(* IEC 61131-3 sources: s7-to-codesys/s7conv/tests/snapshots/fixtures/src/POUs/FB_Legacy, 2 files *)

(* ---- FB_Legacy.decl.st ---- *)
// Назначение: Функциональный блок «FB_Legacy», сконвертирован из SCL
// Автор:      не указан (исходный блок S7); перевод в ST — s7conv 0.1.0
// Версия:     0.1 (исходный блок S7)
// Документ:   docs/CONVERSION_REPORT.md, docs/MAPPING.md
// Источник:   s7conv/tests/fixtures/unsupported.scl, строки 2–44, FUNCTION_BLOCK "FB_Legacy"
// Сгенерировано s7conv: пометки MIGRATION-CHECK и MIGRATION-TODO требуют ручного разбора.
// MIGRATION-CHECK: стандартный (неоптимизированный) доступ S7: абсолютная адресация и порядок байтов не переносятся
//                  (стр. 2)
// MIGRATION-CHECK: реманентность задаётся в экземпляре DB (DB_SPECIFIC) — объявлено VAR (стр. 19)
// ---- комментарий в начале исходного файла SCL ----
// Фикстура s7conv: конструкции, которые конвертер не переводит или переводит с пометкой.
FUNCTION_BLOCK FB_Legacy
VAR_INPUT
    // MIGRATION-TODO: Variant — нет аналога в CODESYS; переписать (ANY, POINTER или перегрузка) (стр. 6)
    // anyIn : Variant;
    // MIGRATION-TODO: DTL — структура S7 (YEAR, MONTH, ...), в CODESYS нет; заменить на DT или свою структуру (стр.
    //                 7)
    // stamp : DTL;
    // MIGRATION-CHECK: имя «time» переименовано в «time_» (ключевое слово CODESYS или повтор) (стр. 8)
    time_ : TIME;
END_VAR
VAR
    raw : WORD;
    // MIGRATION-TODO: AT (наложение переменных S7) — переписать через UNION или битовый доступ (стр. 12)
    // bits AT raw : Array[0..15] of Bool;
    // MIGRATION-CHECK: счётчик S7 → CTU (CODESYS Standard): PV и CV — WORD (0…65535), в S7 — тип счётчика;
    //                  проверить диапазон (стр. 13)
    counter : CTU;
    txt : WSTRING(10);
    // MIGRATION-CHECK: Char → STRING(1): в CODESYS нет типа CHAR, сравнения и CHAR_TO_* проверить (стр. 15)
    ch : STRING(1);
    flags : BYTE;
    // MIGRATION-TODO: TONR (таймер с накоплением) — в CODESYS Standard нет (стр. 17)
    // acc : TONR_TIME;
END_VAR
VAR
    keep : INT;
END_VAR

(* ---- FB_Legacy.impl.st ---- *)
counter(CU := raw.0, RESET := raw.1, PV := 10);
IF counter.Q THEN
    // MIGRATION-TODO: GOTO — переходы не переносятся (переписать структурно) (стр. 26)
    // GOTO done;
    ; // нет операторов
END_IF
// MIGRATION-TODO: PEEK_WORD: нет прямого аналога в CODESYS Standard (стр. 28)
// #raw := PEEK_WORD(area := 16#84, dbNumber := 1, byteOffset := 0);
// MIGRATION-CHECK: срез .%B1 → WORD_TO_BYTE(SHR(...)): нумерация срезов S7 от младшей части — сверить с источником
//                  (стр. 29)
flags := WORD_TO_BYTE(SHR(raw, 8));
// MIGRATION-TODO: оператор не разобран: ожидалось ';', найдено 'ENO' (стр. 30)
// #keep := #keep + 1 ENO => #ok;
txt := "abc";
ch := 'A';
// MIGRATION-CHECK: ROUND → REAL_TO_DINT: правило округления половины (x.5) сверить с источником (стр. 33)
keep := REAL_TO_DINT(2.5) + TRUNC(1.5);
// MIGRATION-TODO: адрес %DB1.DBX0.0 не поддерживается (только %I, %Q, %M) (стр. 34)
// %DB1.DBX0.0 := TRUE;
// MIGRATION-CHECK: отрицательный TIME: в CODESYS TIME беззнаковый (UDINT мс) (стр. 35)
time_ := T#-5s;
raw := SHL(raw, 2) OR WORD#16#00FF;
keep := LIMIT(0, keep, 100);
keep := MAX(1, 2, 3);
// MIGRATION-CHECK: REAL_TO_DWORD: в S7-1200/1500 переносится битовый образ, в CODESYS — числовое значение (стр. 39)
raw := DWORD_TO_WORD(REAL_TO_DWORD(1.0));
// MIGRATION-CHECK: ** → EXPT: тип результата для целых операндов сверить (в S7 — REAL/LREAL) (стр. 40)
keep := EXPT(keep, 2);
// MIGRATION-TODO: метка перехода — переходы не переносятся (стр. 41)
// done:
keep := 0;
// MIGRATION-TODO: DB "Unknown_DB" не найден в корпусе — добавьте его исходник (стр. 42)
// "Unknown_DB".value := 1;
// MIGRATION-TODO: оператор не разобран: ожидалось выражение, найдено ':=' (стр. 43)
// #keep := := 2;
